Staubli VAL3: movePoint.pgx

program movePoint(num x_nStep, num x_nIndex)
  local bool l_bResult
begin
  //   l_bResult=userPageConfirm("是否移动到该点位？")
  //  if l_bResult
  resetMotion()
  $jogMode(0)
  switch x_nStep
    case 0
      movel(savedata:fFrameItem[x_nIndex].pPointRx[0],tUsingTool,mNomSpeed)
    break
    case 1
      movel(savedata:fFrameItem[x_nIndex].pPointRx[1],tUsingTool,mNomSpeed)
    break
    case 2
      movel(savedata:fFrameItem[x_nIndex].pPointRx[2],tUsingTool,mNomSpeed)
    break
  endSwitch
  //  endIf
end
